(* Logix 5000 project; controller R400_500_XLS vendor 1 type 14 code 216 rev 31.11; software revision 31.01; part 8 of 32 *)
(* tags used below, declared in another part *)
   Abort1 : DINT;   // Not Used
   Alarm : SINT;   // Wait 3 seconds
   Ashutdown : SINT;   // Not Used
   bAlrm : BOOL[64];
   Critical_Alarm : BOOL;
   CycExcBuffer : UDT_CYCLE;
   CycleNotEmpty : SINT;
   CycleSequence : UDT_CYCLE_SEQUENCE;
   CycViewBuffer : UDT_WASH;
   DRYING : DINT;   // Drying id number
   FINAL_RINSE_MAX_NBR : INT;   // Maximum nimber of final rinse
   iBuffer : DINT[5];
   InjMan : SINT;
   M : DINT[5];   // Memory Bits
   OneShot : DINT[1];
   ONS_FC34 : DINT;
   PWR_UP : DINT;
   Run : DINT;
   Shutdown : SINT;   // Shutdown sequence steps
   sPrntArray : STRING[300];   // Printer String Array
   Tmr : TIMER[107];
   washerMode : SINT;   // Washer Mode Flag 0 -> Ready; 1 -> Supervisor; 2 -> Service; 3 -> Run.
   AlarmTrigger : INT;   // Triggers the alarm screen if different of 0
   bAcceptRejectRecorded : BOOL;   // Cycle Accept/Reject Recorded By User
   bHMICycleAccepted : BOOL;   // HMI - Button Cycle Accepted
   bHMICycleRejected : BOOL;   // HMI - Button Cycle Rejected
   bONSCycleAccepted : BOOL;
   bONSCycleRejected : BOOL;
   Current_Screen : DINT;
   CurrentUser : STRING;   // Current User
   Doors_Check : DINT;
   I_Ld_Dr_Cls_Sw : BOOL;   // Load door close
   I_Ld_Dr_Obs_Sw : BOOL;   // Load door obstruction switch
   I_Unld_Dr_Cls_Sw : BOOL;   // Unload door close
   I_Unld_Dr_Obs_Sw : BOOL;   // Unload door obstruction switch
   I_UnldDr_ClseSlnce_Bttn : BOOL;   // Door Close/ Silence button Unload Side
   I_UnldDr_Opn_Bttn : BOOL;   // Door Open button Unload side
   Load : Doors;
   LoadDoorClosing : BOOL;
   LoadDoorOpening : BOOL;
   MaintainCloseLd : BOOL;
   MaintainCloseUnld : BOOL;
   MaintainOpenLd : BOOL;
   MaintainOpenUnld : BOOL;
   Msg_Door : SINT;   // 1= Door(s) not closed
   Msg_DoorSteps : INT;   // Display Safety Door Test Messages
   Msg_TempSp : SINT;   // HMI Information Message tag
   previous_s108 : DINT;
   PrintIndex : DINT;
   Q_Ld_Dr_Clse_Vlv : BOOL;   // Load door close pilot valve
   Q_Ld_Dr_Opn_Vlv : BOOL;   // Load door open pilot valve
   Q_Unld_Dr_Clse_Vlve : BOOL;   // Unload door close pilot valve
   Q_Unld_Dr_Opn_Vlve : BOOL;   // Unload door open pilot valve
   Screen_Ctrl : DINT;   // PLC Screen Request
   sCycleAccepted : STRING;   // Cycle Accepted
   sCycleRejected : STRING;   // Cycle Rejected
   Selector : UDT_SELECTOR[25];   // Piloted list selector
   SelectorView : UDT_SELECTOR[3];   // Piloted list selector for cycle view menu
   Tpb : DINT[11];
   TpbImage : DINT[11];
   Unit : Hrdwre;   // Unit Configuration
   UnLoad : Doors;
   UnloadDoorClosing : BOOL;
   UnloadDoorOpening : BOOL;
(* MainProgram, continued *)

ROUTINE OPR_1_WSH_11_14_OPN_CLSD_LD_DR   (* ladder *)
// Module to open or close the Load door
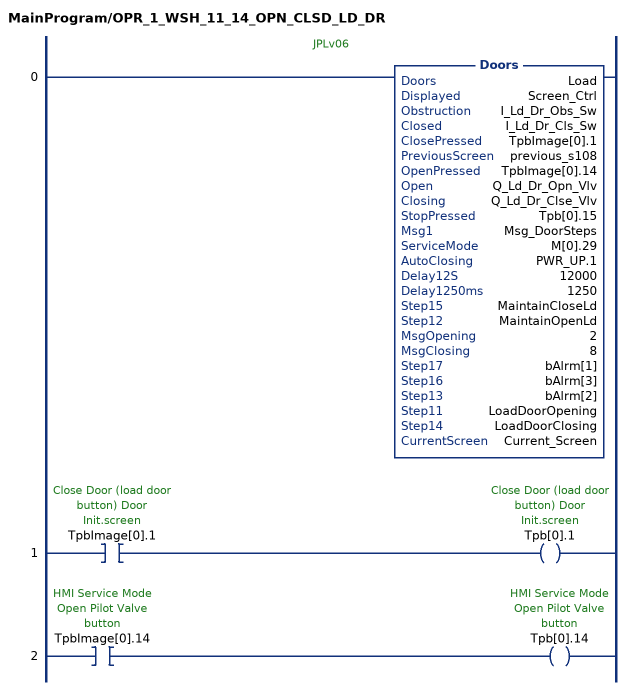
   // JPLv06
   0: Doors(Load,Screen_Ctrl,I_Ld_Dr_Obs_Sw,I_Ld_Dr_Cls_Sw,TpbImage[0].1,previous_s108,TpbImage[0].14,Q_Ld_Dr_Opn_Vlv,Q_Ld_Dr_Clse_Vlv,Tpb[0].15,Msg_DoorSteps,M[0].29,PWR_UP.1,12000,1250,MaintainCloseLd,MaintainOpenLd,2,8,bAlrm[1],bAlrm[3],bAlrm[2],LoadDoorOpening,LoadDoorClosing,Current_Screen);
   1: XIC(TpbImage[0].1)OTE(Tpb[0].1);
   2: XIC(TpbImage[0].14)OTE(Tpb[0].14);
END_ROUTINE

ROUTINE OPR_1_WSH_11_14_OPN_CLSD_UNLD_DR   (* ladder *)
// Module to open or close the unload door
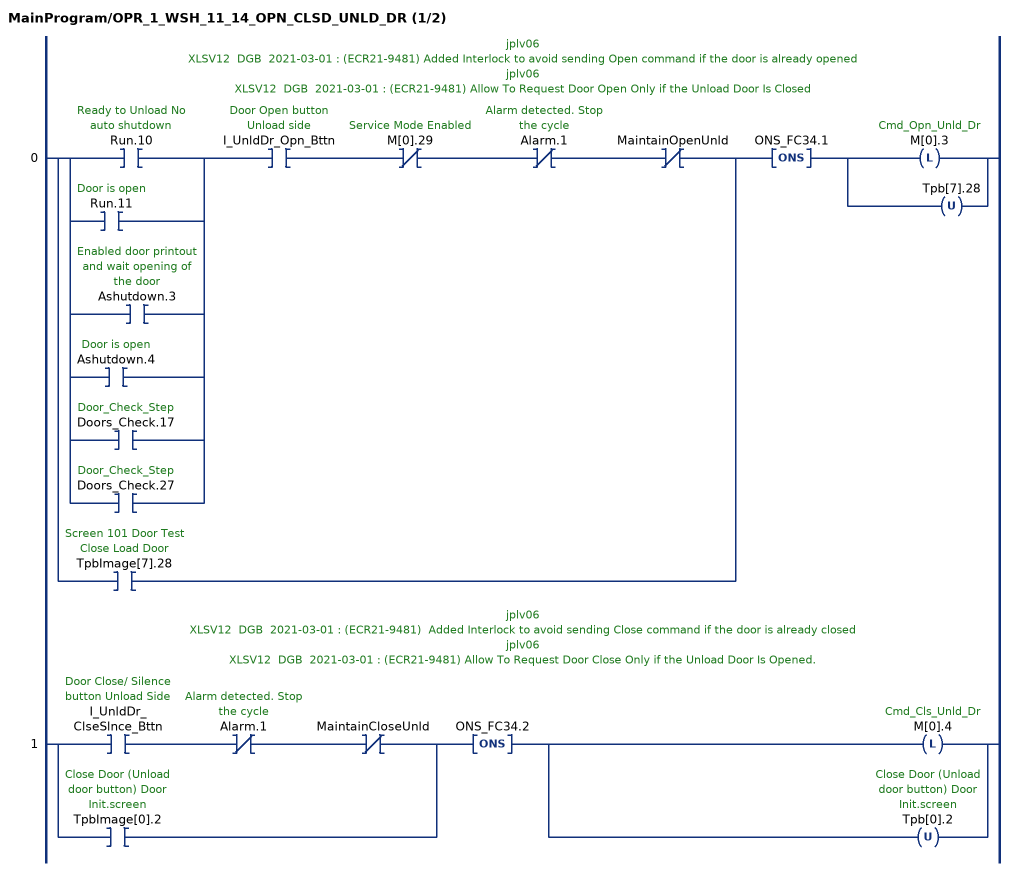
   // jplv06
   // XLSV12  DGB  2021-03-01 : (ECR21-9481) Added Interlock to avoid sending Open command if the door is already opened
   // jplv06
   // XLSV12  DGB  2021-03-01 : (ECR21-9481) Allow To Request Door Open Only if the Unload Door Is Closed
   0: [[XIC(Run.10) ,XIC(Run.11) ,XIC(Ashutdown.3) ,XIC(Ashutdown.4) ,XIC(Doors_Check.17) ,XIC(Doors_Check.27) ] XIC(I_UnldDr_Opn_Bttn) XIO(M[0].29) XIO(Alarm.1) XIO(MaintainOpenUnld) ,XIC(TpbImage[7].28) ]ONS(ONS_FC34.1)[OTL(M[0].3) ,OTU(Tpb[7].28) ];
   // jplv06
   // XLSV12  DGB  2021-03-01 : (ECR21-9481)  Added Interlock to avoid sending Close command if the door is already closed
   // jplv06
   // XLSV12  DGB  2021-03-01 : (ECR21-9481) Allow To Request Door Close Only if the Unload Door Is Opened.
   1: [XIC(I_UnldDr_ClseSlnce_Bttn) XIO(Alarm.1) XIO(MaintainCloseUnld) ,XIC(TpbImage[0].2) ]ONS(ONS_FC34.2)[OTL(M[0].4) ,OTU(Tpb[0].2) ];
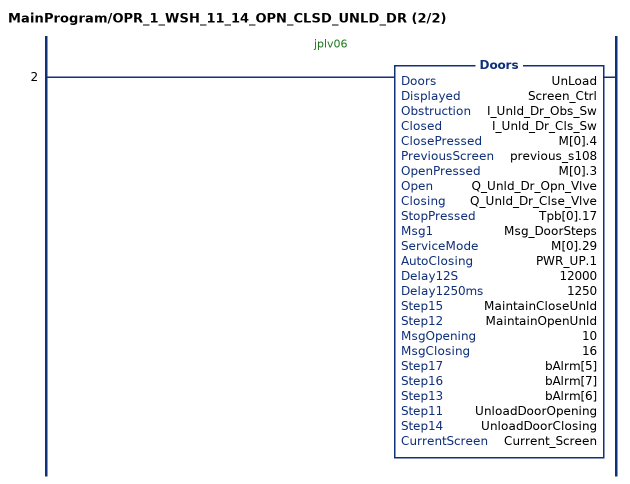
   // jplv06
   2: Doors(UnLoad,Screen_Ctrl,I_Unld_Dr_Obs_Sw,I_Unld_Dr_Cls_Sw,M[0].4,previous_s108,M[0].3,Q_Unld_Dr_Opn_Vlve,Q_Unld_Dr_Clse_Vlve,Tpb[0].17,Msg_DoorSteps,M[0].29,PWR_UP.1,12000,1250,MaintainCloseUnld,MaintainOpenUnld,10,16,bAlrm[5],bAlrm[7],bAlrm[6],UnloadDoorOpening,UnloadDoorClosing,Current_Screen);
END_ROUTINE

ROUTINE OPR_2_OPR_3_OPR_4_VIEW_CYCLE   (* ladder *)
// This routine manages the HMI screens in order for the operator to view the cycle parameters
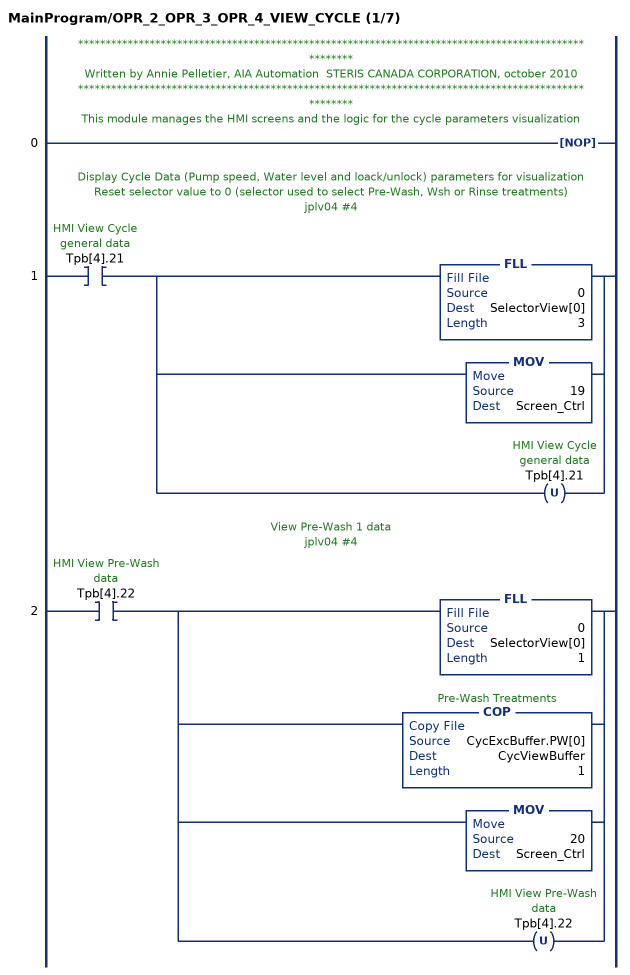
   // ****************************************************************************************************
   // Written by Annie Pelletier, AIA Automation  STERIS CANADA CORPORATION, october 2010
   // ****************************************************************************************************
   // This module manages the HMI screens and the logic for the cycle parameters visualization
   0: NOP();
   // Display Cycle Data (Pump speed, Water level and loack/unlock) parameters for visualization
   // Reset selector value to 0 (selector used to select Pre-Wash, Wsh or Rinse treatments)
   // jplv04 #4
   1: XIC(Tpb[4].21)[FLL(0,SelectorView[0],3) ,MOV(19,Screen_Ctrl) ,OTU(Tpb[4].21) ];
   // View Pre-Wash 1 data
   // jplv04 #4
   2: XIC(Tpb[4].22)[FLL(0,SelectorView[0],1) ,COP(CycExcBuffer.PW[0],CycViewBuffer,1) ,MOV(20,Screen_Ctrl) ,OTU(Tpb[4].22) ];
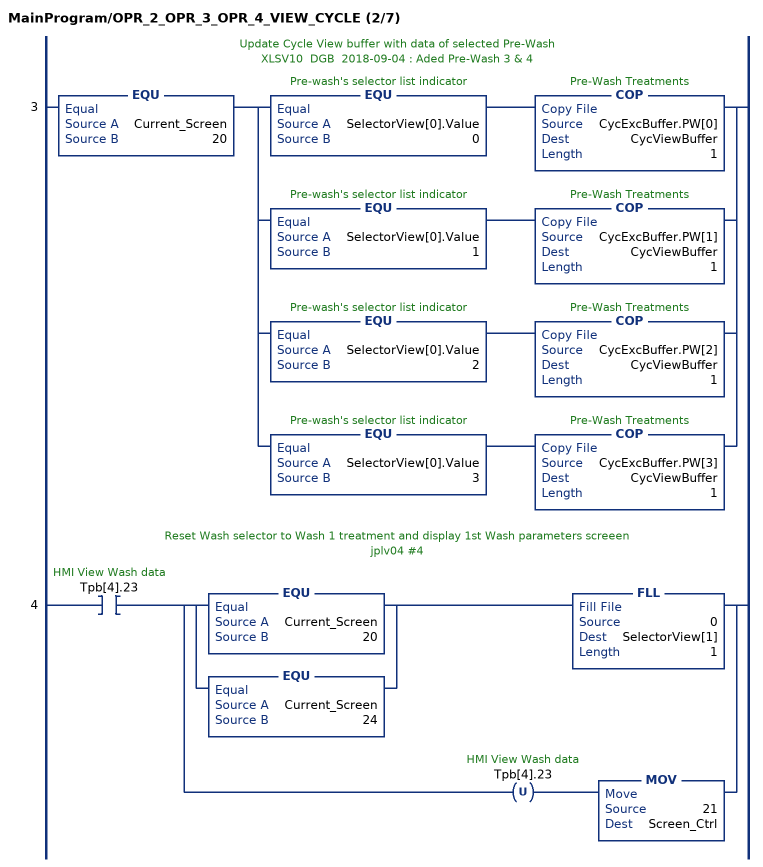
   // Update Cycle View buffer with data of selected Pre-Wash
   // XLSV10  DGB  2018-09-04 : Aded Pre-Wash 3 & 4
   3: EQU(Current_Screen,20)[EQU(SelectorView[0].Value,0) COP(CycExcBuffer.PW[0],CycViewBuffer,1) ,EQU(SelectorView[0].Value,1) COP(CycExcBuffer.PW[1],CycViewBuffer,1) ,EQU(SelectorView[0].Value,2) COP(CycExcBuffer.PW[2],CycViewBuffer,1) ,EQU(SelectorView[0].Value,3) COP(CycExcBuffer.PW[3],CycViewBuffer,1) ];
   // Reset Wash selector to Wash 1 treatment and display 1st Wash parameters screeen
   // jplv04 #4
   4: XIC(Tpb[4].23)[[EQU(Current_Screen,20) ,EQU(Current_Screen,24) ] FLL(0,SelectorView[1],1) ,OTU(Tpb[4].23) MOV(21,Screen_Ctrl) ];
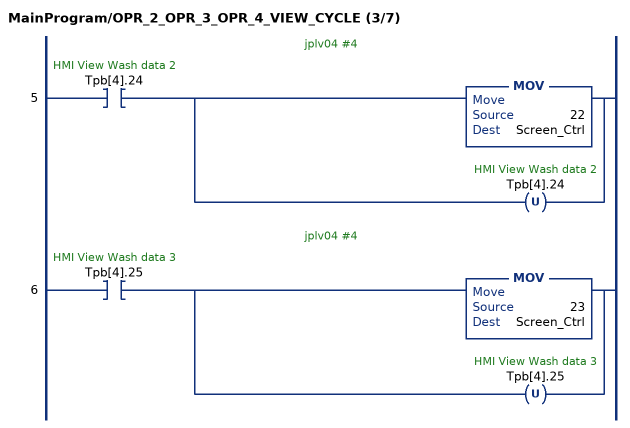
   // jplv04 #4
   5: XIC(Tpb[4].24)[MOV(22,Screen_Ctrl) ,OTU(Tpb[4].24) ];
   // jplv04 #4
   6: XIC(Tpb[4].25)[MOV(23,Screen_Ctrl) ,OTU(Tpb[4].25) ];
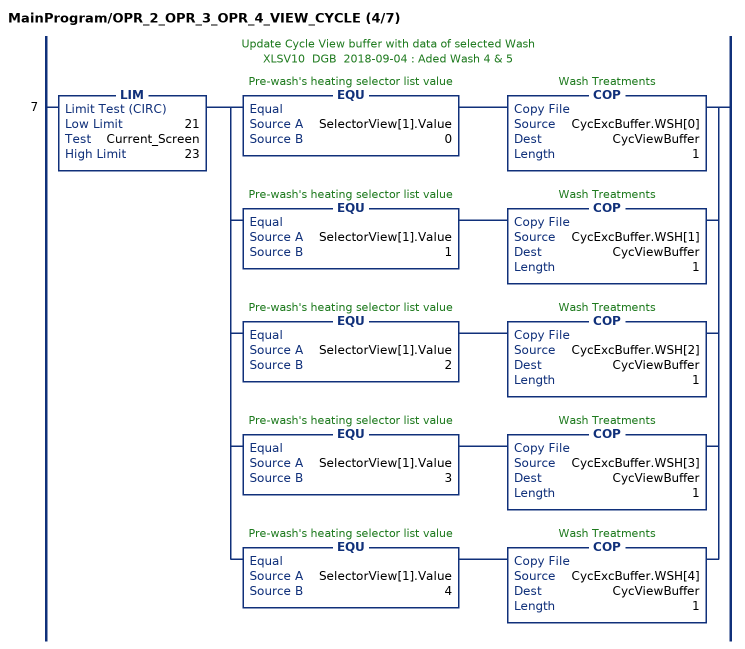
   // Update Cycle View buffer with data of selected Wash
   // XLSV10  DGB  2018-09-04 : Aded Wash 4 & 5
   7: LIM(21,Current_Screen,23)[EQU(SelectorView[1].Value,0) COP(CycExcBuffer.WSH[0],CycViewBuffer,1) ,EQU(SelectorView[1].Value,1) COP(CycExcBuffer.WSH[1],CycViewBuffer,1) ,EQU(SelectorView[1].Value,2) COP(CycExcBuffer.WSH[2],CycViewBuffer,1) ,EQU(SelectorView[1].Value,3) COP(CycExcBuffer.WSH[3],CycViewBuffer,1) ,EQU(SelectorView[1].Value,4) COP(CycExcBuffer.WSH[4],CycViewBuffer,1) ];
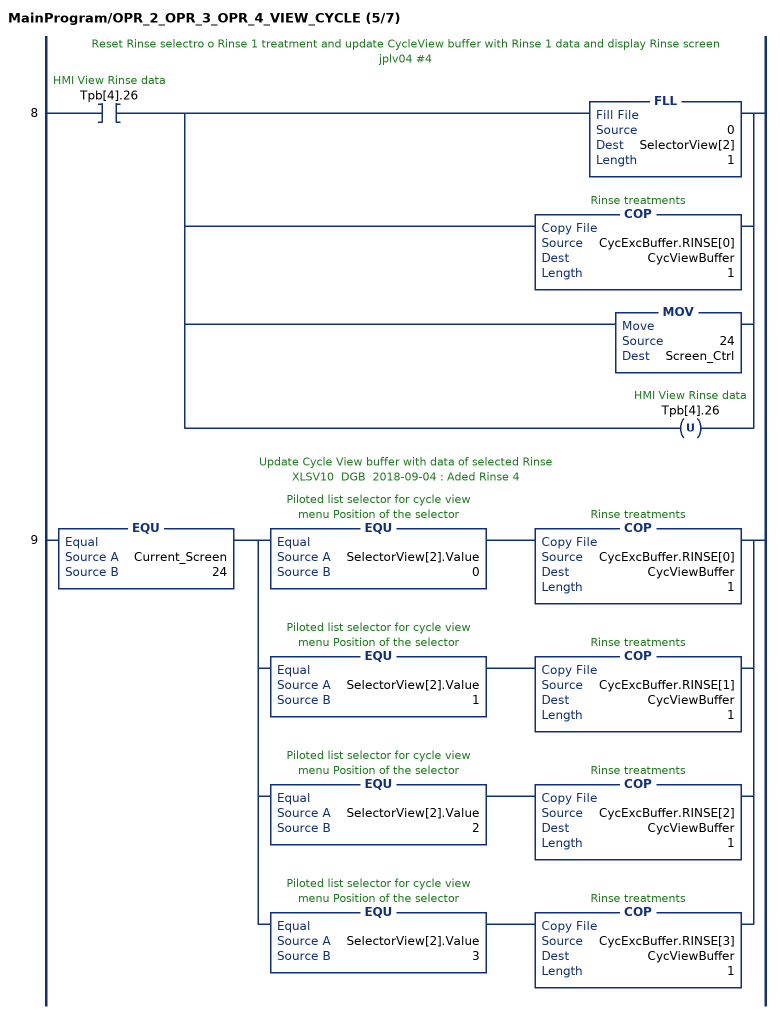
   // Reset Rinse selectro o Rinse 1 treatment and update CycleView buffer with Rinse 1 data and display Rinse screen
   // jplv04 #4
   8: XIC(Tpb[4].26)[FLL(0,SelectorView[2],1) ,COP(CycExcBuffer.RINSE[0],CycViewBuffer,1) ,MOV(24,Screen_Ctrl) ,OTU(Tpb[4].26) ];
   // Update Cycle View buffer with data of selected Rinse
   // XLSV10  DGB  2018-09-04 : Aded Rinse 4
   9: EQU(Current_Screen,24)[EQU(SelectorView[2].Value,0) COP(CycExcBuffer.RINSE[0],CycViewBuffer,1) ,EQU(SelectorView[2].Value,1) COP(CycExcBuffer.RINSE[1],CycViewBuffer,1) ,EQU(SelectorView[2].Value,2) COP(CycExcBuffer.RINSE[2],CycViewBuffer,1) ,EQU(SelectorView[2].Value,3) COP(CycExcBuffer.RINSE[3],CycViewBuffer,1) ];
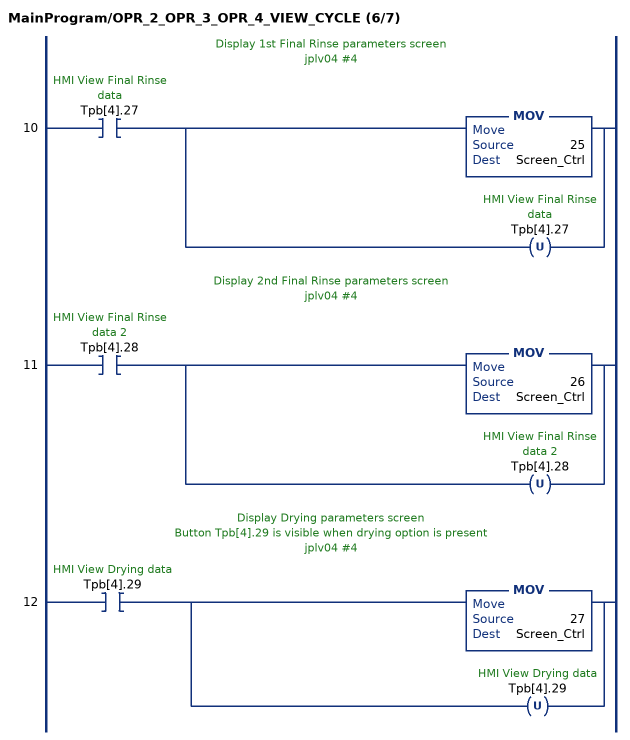
   // Display 1st Final Rinse parameters screen
   // jplv04 #4
   10: XIC(Tpb[4].27)[MOV(25,Screen_Ctrl) ,OTU(Tpb[4].27) ];
   // Display 2nd Final Rinse parameters screen
   // jplv04 #4
   11: XIC(Tpb[4].28)[MOV(26,Screen_Ctrl) ,OTU(Tpb[4].28) ];
   // Display Drying parameters screen
   // Button Tpb[4].29 is visible when drying option is present
   // jplv04 #4
   12: XIC(Tpb[4].29)[MOV(27,Screen_Ctrl) ,OTU(Tpb[4].29) ];
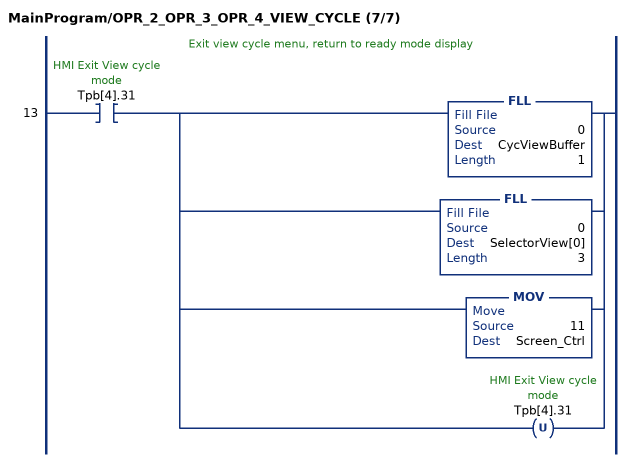
   // Exit view cycle menu, return to ready mode display
   13: XIC(Tpb[4].31)[FLL(0,CycViewBuffer,1) ,FLL(0,SelectorView[0],3) ,MOV(11,Screen_Ctrl) ,OTU(Tpb[4].31) ];
END_ROUTINE

ROUTINE OPR_8_OPR_11_WSH_58_RUN_PAUSE_CMPLTE_CYC   (* ladder *)
// This module start the cycle and manage the stop/resume function
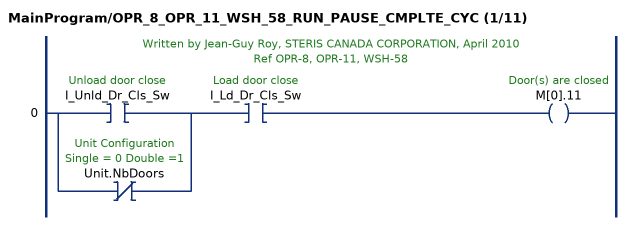
   // Written by Jean-Guy Roy, STERIS CANADA CORPORATION, April 2010
   // Ref OPR-8, OPR-11, WSH-58
   0: [XIC(I_Unld_Dr_Cls_Sw) ,XIO(Unit.NbDoors) ]XIC(I_Ld_Dr_Cls_Sw)OTE(M[0].11);
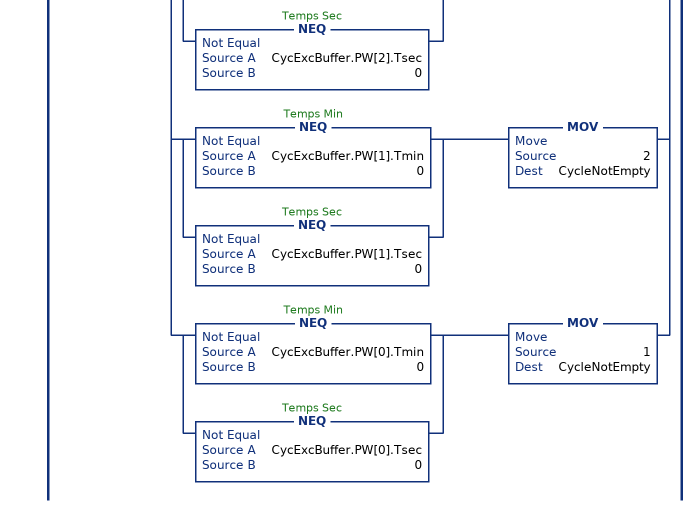
   // When start button is pressed, this rung checks if a recirculated treatment is present in the cycle
   // Check Rinse 3 Treatment time
   // jplv04 #4
   // XLSV10  DGB  2018-09-17 : Added To support New Treatment
   1: XIC(TpbImage[0].3)[[NEQ(CycExcBuffer.RINSE[3].Tmin,0) ,NEQ(CycExcBuffer.RINSE[3].Tsec,0) ] MOV(13,CycleNotEmpty) ,[NEQ(CycExcBuffer.RINSE[2].Tmin,0) ,NEQ(CycExcBuffer.RINSE[2].Tsec,0) ] MOV(12,CycleNotEmpty) ,[NEQ(CycExcBuffer.RINSE[1].Tmin,0) ,NEQ(CycExcBuffer.RINSE[1].Tsec,0) ] MOV(11,CycleNotEmpty) ,[NEQ(CycExcBuffer.RINSE[0].Tmin,0) ,NEQ(CycExcBuffer.RINSE[0].Tsec,0) ] MOV(10,CycleNotEmpty) ,[NEQ(CycExcBuffer.WSH[4].Tmin,0) ,NEQ(CycExcBuffer.WSH[4].Tsec,0) ] MOV(9,CycleNotEmpty) ,[NEQ(CycExcBuffer.WSH[3].Tmin,0) ,NEQ(CycExcBuffer.WSH[3].Tsec,0) ] MOV(8,CycleNotEmpty) ,[NEQ(CycExcBuffer.WSH[2].Tmin,0) ,NEQ(CycExcBuffer.WSH[2].Tsec,0) ] MOV(7,CycleNotEmpty) ,[NEQ(CycExcBuffer.WSH[1].Tmin,0) ,NEQ(CycExcBuffer.WSH[1].Tsec,0) ] MOV(6,CycleNotEmpty) ,[NEQ(CycExcBuffer.WSH[0].Tmin,0) ,NEQ(CycExcBuffer.WSH[0].Tsec,0) ] MOV(5,CycleNotEmpty) ,[NEQ(CycExcBuffer.PW[3].Tmin,0) ,NEQ(CycExcBuffer.PW[3].Tsec,0) ] MOV(4,CycleNotEmpty) ,[NEQ(CycExcBuffer.PW[2].Tmin,0) ,NEQ(CycExcBuffer.PW[2].Tsec,0) ] MOV(3,CycleNotEmpty) ,[NEQ(CycExcBuffer.PW[1].Tmin,0) ,NEQ(CycExcBuffer.PW[1].Tsec,0) ] MOV(2,CycleNotEmpty) ,[NEQ(CycExcBuffer.PW[0].Tmin,0) ,NEQ(CycExcBuffer.PW[0].Tsec,0) ] MOV(1,CycleNotEmpty) ];
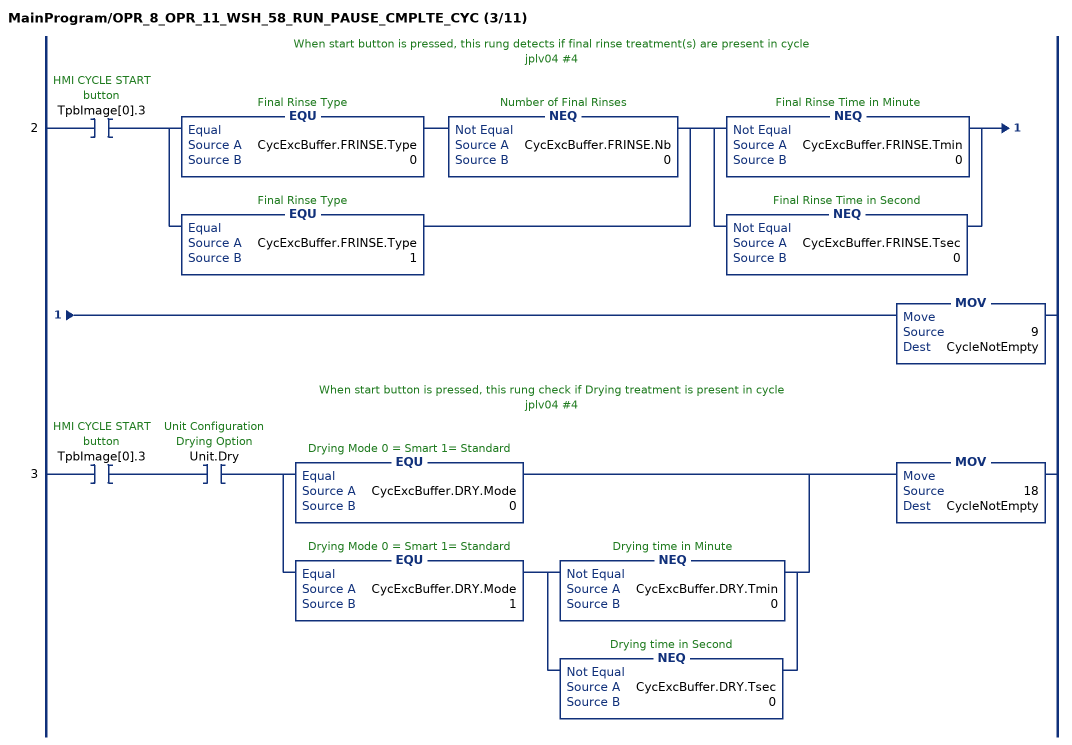
   // When start button is pressed, this rung detects if final rinse treatment(s) are present in cycle
   // jplv04 #4
   2: XIC(TpbImage[0].3)[EQU(CycExcBuffer.FRINSE.Type,0) NEQ(CycExcBuffer.FRINSE.Nb,0) ,EQU(CycExcBuffer.FRINSE.Type,1) ][NEQ(CycExcBuffer.FRINSE.Tmin,0) ,NEQ(CycExcBuffer.FRINSE.Tsec,0) ]MOV(9,CycleNotEmpty);
   // When start button is pressed, this rung check if Drying treatment is present in cycle
   // jplv04 #4
   3: XIC(TpbImage[0].3)XIC(Unit.Dry)[EQU(CycExcBuffer.DRY.Mode,0) ,EQU(CycExcBuffer.DRY.Mode,1) [NEQ(CycExcBuffer.DRY.Tmin,0) ,NEQ(CycExcBuffer.DRY.Tsec,0) ] ]MOV(18,CycleNotEmpty);
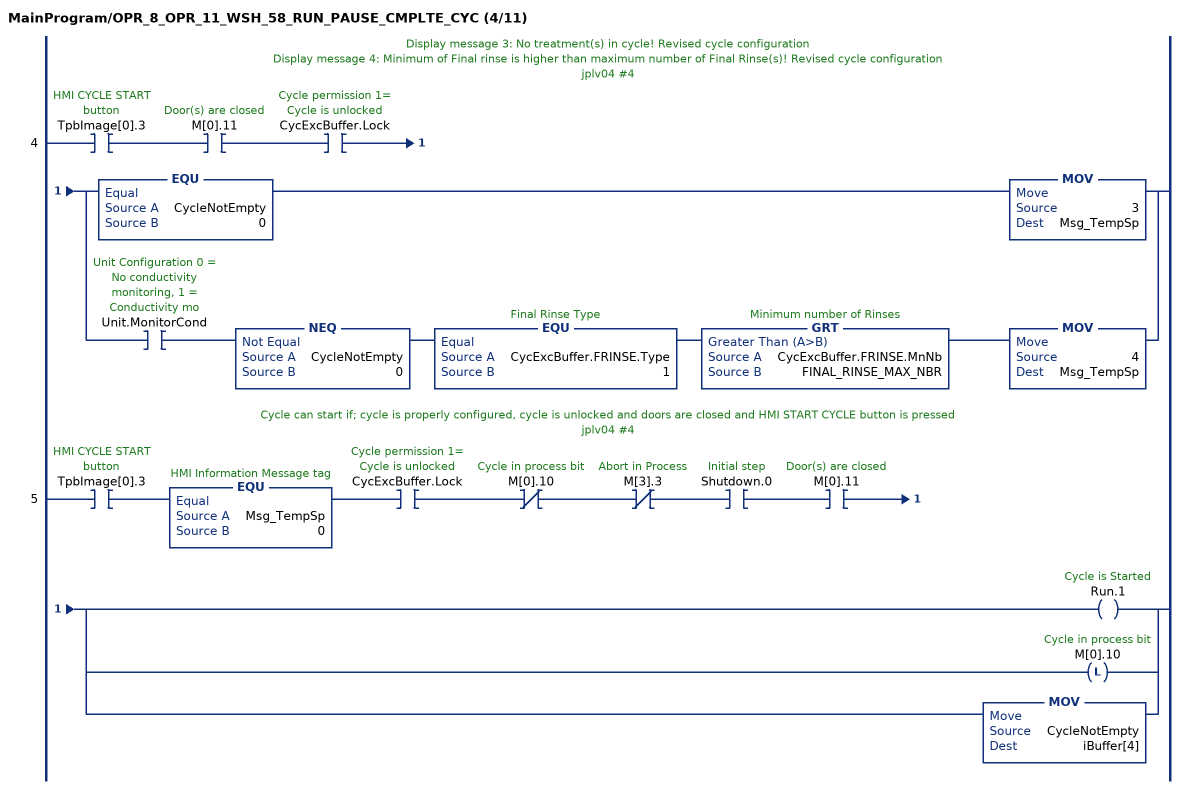
   // Display message 3: No treatment(s) in cycle! Revised cycle configuration
   // Display message 4: Minimum of Final rinse is higher than maximum number of Final Rinse(s)! Revised cycle configuration
   // jplv04 #4
   4: XIC(TpbImage[0].3)XIC(M[0].11)XIC(CycExcBuffer.Lock)[EQU(CycleNotEmpty,0) MOV(3,Msg_TempSp) ,XIC(Unit.MonitorCond) NEQ(CycleNotEmpty,0) EQU(CycExcBuffer.FRINSE.Type,1) GRT(CycExcBuffer.FRINSE.MnNb,FINAL_RINSE_MAX_NBR) MOV(4,Msg_TempSp) ];
   // Cycle can start if; cycle is properly configured, cycle is unlocked and doors are closed and HMI START CYCLE button is pressed
   // jplv04 #4
   5: XIC(TpbImage[0].3)EQU(Msg_TempSp,0)XIC(CycExcBuffer.Lock)XIO(M[0].10)XIO(M[3].3)XIC(Shutdown.0)XIC(M[0].11)[OTE(Run.1) ,OTL(M[0].10) ,MOV(CycleNotEmpty,iBuffer[4]) ];
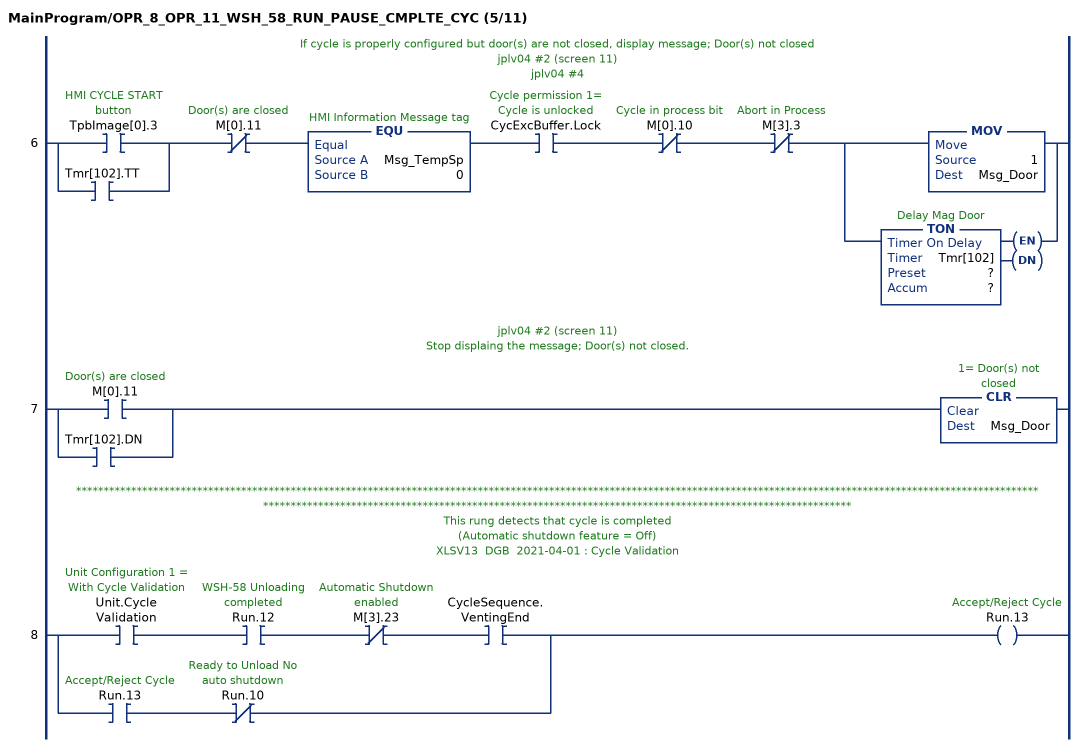
   // If cycle is properly configured but door(s) are not closed, display message; Door(s) not closed
   // jplv04 #2 (screen 11)
   // jplv04 #4
   6: [XIC(TpbImage[0].3) ,XIC(Tmr[102].TT) ]XIO(M[0].11)EQU(Msg_TempSp,0)XIC(CycExcBuffer.Lock)XIO(M[0].10)XIO(M[3].3)[MOV(1,Msg_Door) ,TON(Tmr[102],?,?) ];
   // jplv04 #2 (screen 11)
   // Stop displaing the message; Door(s) not closed.
   7: [XIC(M[0].11) ,XIC(Tmr[102].DN) ]CLR(Msg_Door);
   // ******************************************************************************************************************************************************************************************************************************************************************************************
   // This rung detects that cycle is completed
   // (Automatic shutdown feature = Off)
   // XLSV13  DGB  2021-04-01 : Cycle Validation
   8: [XIC(Unit.CycleValidation) XIC(Run.12) XIO(M[3].23) XIC(CycleSequence.VentingEnd) ,XIC(Run.13) XIO(Run.10) ]OTE(Run.13);
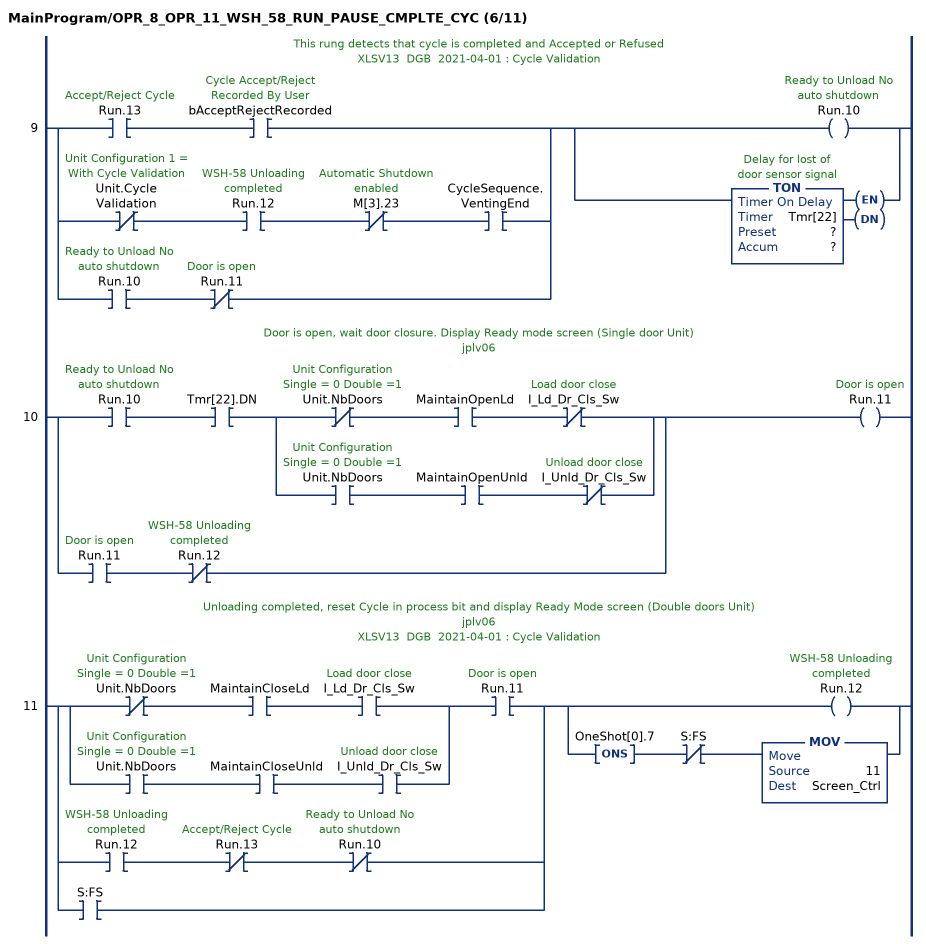
   // This rung detects that cycle is completed and Accepted or Refused
   // XLSV13  DGB  2021-04-01 : Cycle Validation
   9: [XIC(Run.13) XIC(bAcceptRejectRecorded) ,XIO(Unit.CycleValidation) XIC(Run.12) XIO(M[3].23) XIC(CycleSequence.VentingEnd) ,XIC(Run.10) XIO(Run.11) ][OTE(Run.10) ,TON(Tmr[22],?,?) ];
   // Door is open, wait door closure. Display Ready mode screen (Single door Unit)
   // jplv06
   10: [XIC(Run.10) XIC(Tmr[22].DN) [XIO(Unit.NbDoors) XIC(MaintainOpenLd) XIO(I_Ld_Dr_Cls_Sw) ,XIC(Unit.NbDoors) XIC(MaintainOpenUnld) XIO(I_Unld_Dr_Cls_Sw) ] ,XIC(Run.11) XIO(Run.12) ]OTE(Run.11);
   // Unloading completed, reset Cycle in process bit and display Ready Mode screen (Double doors Unit)
   // jplv06
   // XLSV13  DGB  2021-04-01 : Cycle Validation
   11: [[XIO(Unit.NbDoors) XIC(MaintainCloseLd) XIC(I_Ld_Dr_Cls_Sw) ,XIC(Unit.NbDoors) XIC(MaintainCloseUnld) XIC(I_Unld_Dr_Cls_Sw) ] XIC(Run.11) ,XIC(Run.12) XIO(Run.13) XIO(Run.10) ,XIC(S:FS) ][OTE(Run.12) ,ONS(OneShot[0].7) XIO(S:FS) MOV(11,Screen_Ctrl) ];
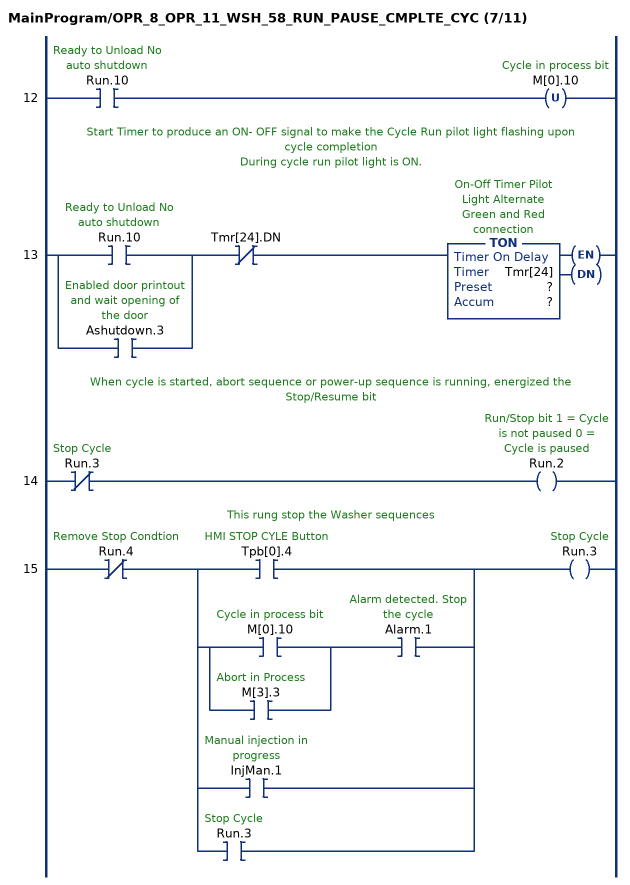
   12: XIC(Run.10)OTU(M[0].10);
   // Start Timer to produce an ON- OFF signal to make the Cycle Run pilot light flashing upon cycle completion
   // During cycle run pilot light is ON.
   13: [XIC(Run.10) ,XIC(Ashutdown.3) ]XIO(Tmr[24].DN)TON(Tmr[24],?,?);
   // When cycle is started, abort sequence or power-up sequence is running, energized the Stop/Resume bit
   14: XIO(Run.3)OTE(Run.2);
   // This rung stop the Washer sequences
   15: XIO(Run.4)[XIC(Tpb[0].4) ,[XIC(M[0].10) ,XIC(M[3].3) ] XIC(Alarm.1) ,XIC(InjMan.1) ,XIC(Run.3) ]OTE(Run.3);
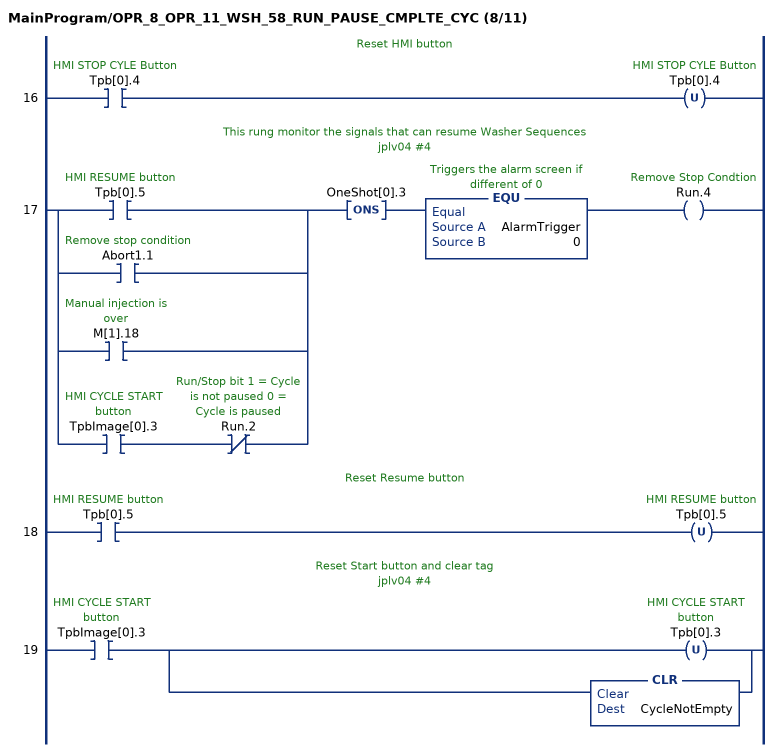
   // Reset HMI button
   16: XIC(Tpb[0].4)OTU(Tpb[0].4);
   // This rung monitor the signals that can resume Washer Sequences
   // jplv04 #4
   17: [XIC(Tpb[0].5) ,XIC(Abort1.1) ,XIC(M[1].18) ,XIC(TpbImage[0].3) XIO(Run.2) ]ONS(OneShot[0].3)EQU(AlarmTrigger,0)OTE(Run.4);
   // Reset Resume button
   18: XIC(Tpb[0].5)OTU(Tpb[0].5);
   // Reset Start button and clear tag
   // jplv04 #4
   19: XIC(TpbImage[0].3)[OTU(Tpb[0].3) ,CLR(CycleNotEmpty) ];
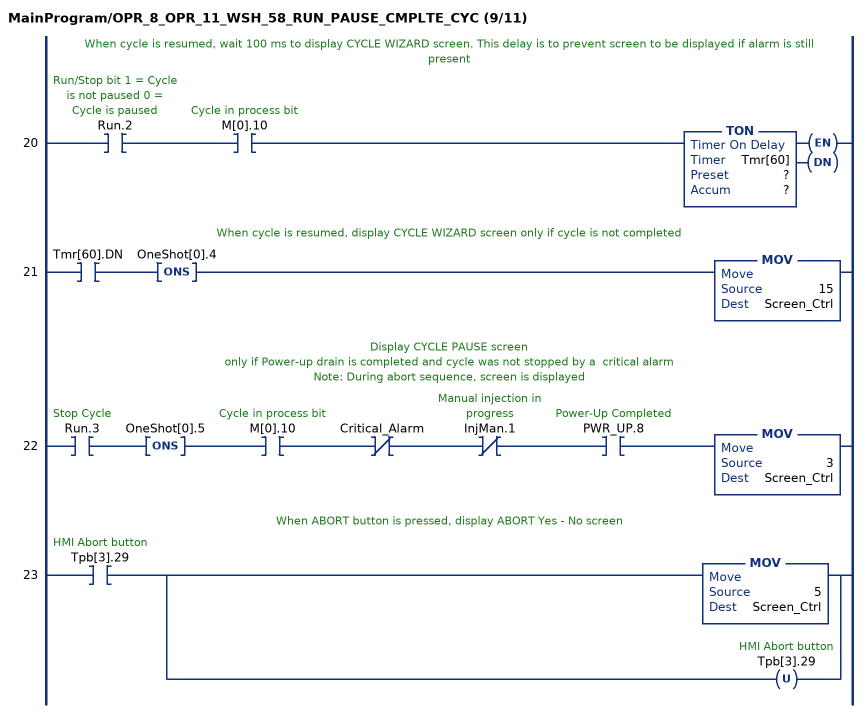
   // When cycle is resumed, wait 100 ms to display CYCLE WIZARD screen. This delay is to prevent screen to be displayed if alarm is still present
   20: XIC(Run.2)XIC(M[0].10)TON(Tmr[60],?,?);
   // When cycle is resumed, display CYCLE WIZARD screen only if cycle is not completed
   21: XIC(Tmr[60].DN)ONS(OneShot[0].4)MOV(15,Screen_Ctrl);
   // Display CYCLE PAUSE screen
   // only if Power-up drain is completed and cycle was not stopped by a  critical alarm
   // Note: During abort sequence, screen is displayed
   22: XIC(Run.3)ONS(OneShot[0].5)XIC(M[0].10)XIO(Critical_Alarm)XIO(InjMan.1)XIC(PWR_UP.8)MOV(3,Screen_Ctrl);
   // When ABORT button is pressed, display ABORT Yes - No screen
   23: XIC(Tpb[3].29)[MOV(5,Screen_Ctrl) ,OTU(Tpb[3].29) ];
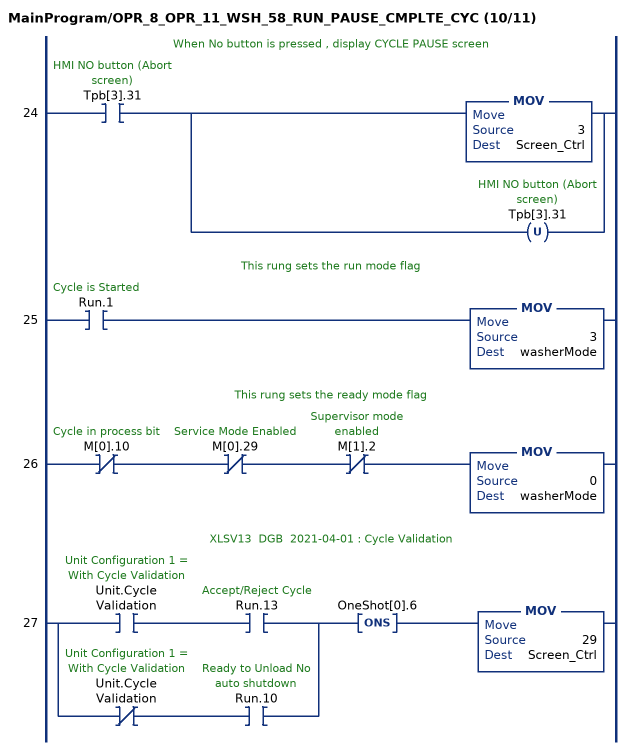
   // When No button is pressed , display CYCLE PAUSE screen
   24: XIC(Tpb[3].31)[MOV(3,Screen_Ctrl) ,OTU(Tpb[3].31) ];
   // This rung sets the run mode flag
   25: XIC(Run.1)MOV(3,washerMode);
   // This rung sets the ready mode flag
   26: XIO(M[0].10)XIO(M[0].29)XIO(M[1].2)MOV(0,washerMode);
   // XLSV13  DGB  2021-04-01 : Cycle Validation
   27: [XIC(Unit.CycleValidation) XIC(Run.13) ,XIO(Unit.CycleValidation) XIC(Run.10) ]ONS(OneShot[0].6)MOV(29,Screen_Ctrl);
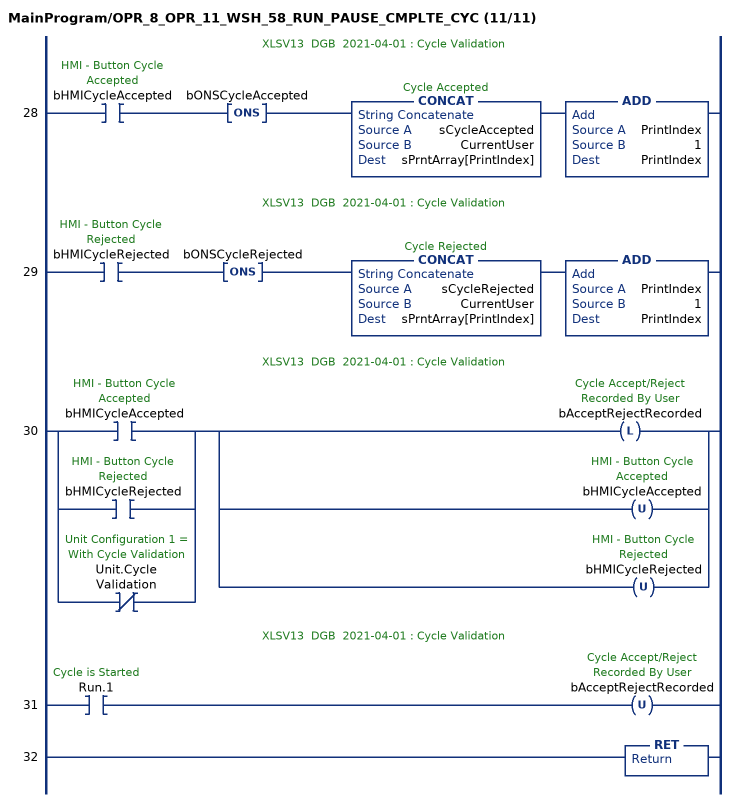
   // XLSV13  DGB  2021-04-01 : Cycle Validation
   28: XIC(bHMICycleAccepted)ONS(bONSCycleAccepted)CONCAT(sCycleAccepted,CurrentUser,sPrntArray[PrintIndex])ADD(PrintIndex,1,PrintIndex);
   // XLSV13  DGB  2021-04-01 : Cycle Validation
   29: XIC(bHMICycleRejected)ONS(bONSCycleRejected)CONCAT(sCycleRejected,CurrentUser,sPrntArray[PrintIndex])ADD(PrintIndex,1,PrintIndex);
   // XLSV13  DGB  2021-04-01 : Cycle Validation
   30: [XIC(bHMICycleAccepted) ,XIC(bHMICycleRejected) ,XIO(Unit.CycleValidation) ][OTL(bAcceptRejectRecorded) ,OTU(bHMICycleAccepted) ,OTU(bHMICycleRejected) ];
   // XLSV13  DGB  2021-04-01 : Cycle Validation
   31: XIC(Run.1)OTU(bAcceptRejectRecorded);
   32: RET();
END_ROUTINE
